SYSTEM ImportExportTestSystem (* System with a device and resource *)
  (* Standard: 61499-1; Description: Copyright (c) 2026 Martin Erich Jobst This program and the accompanying materials are made available under the terms of the Eclipse Public License 2.0 which is available at https://www.eclipse.org/legal/epl-2.0/ SPDX-License-Identifier: EPL-2.0 *)
  (* Version 1.0, 2026-10-23, Martin Jobst *)
  {SET_ATTRIBUTE(IntegerAttribute, 18)}
  APPLICATION TestApplication (* Application using the basic FB *)
    {SET_ATTRIBUTE(IntegerAttribute, 19)}
    (* Application network comment *)
    FBS
      Basic : fixture::basic::BasicTest;
      Composite : CompositeTest;
      Mapped : fixture::basic::BasicTest;
      Mapped2 : fixture::basic::BasicTest;
    END_FBS
    EVENT_CONNECTIONS
      Basic.CNF TO Composite.REQ; (* Application event connection *)
      Mapped.CNF TO Mapped2.REQ; (* Mapped event connection *)
    END_CONNECTIONS
    DATA_CONNECTIONS
      Basic.DO1 TO Composite.DI1; {SET_ATTRIBUTE(Negated, TRUE)}
    END_CONNECTIONS
    ADAPTER_CONNECTIONS
      Basic.EVENT TO Composite.EVENT;
    END_CONNECTIONS
  END_APPLICATION
  DEVICE TestDeviceInstance : TestDevice(DEVICE_ID := DINT#17 {SET_ATTRIBUTE(IntegerAttribute, 21)}) (* Fixture device *)
    {SET_ATTRIBUTE(Profile, FixtureProfile)}
    {SET_ATTRIBUTE(IntegerAttribute, 22)}
    RESOURCE TestResourceInstance : TestResource(RESOURCE_ID := DINT#23) (* Fixture resource *)
      {SET_ATTRIBUTE(IntegerAttribute, 23)}
      FBS
        Processor : fixture::basic::BasicTest;
        Controller : CompositeTest;
      END_FBS
      EVENT_CONNECTIONS
        Processor.CNF TO Controller.REQ; (* Resource event connection *)
      END_CONNECTIONS
      DATA_CONNECTIONS
        Processor.DO1 TO Controller.DI1;
      END_CONNECTIONS
      ADAPTER_CONNECTIONS
        Processor.EVENT TO Controller.EVENT;
      END_CONNECTIONS
    END_RESOURCE
  END_DEVICE
  MAPPINGS
    TestApplication.Mapped ON TestDeviceInstance.TestResourceInstance;
    TestApplication.Mapped2 ON TestDeviceInstance.TestResourceInstance;
  END_MAPPINGS
  SEGMENTS
    TestSegmentInstance : TestSegment; (* Fixture segment *) {SET_ATTRIBUTE(IntegerAttribute, 24)}
  END_SEGMENTS
  LINKS
    TestDeviceInstance => TestSegmentInstance; (* Fixture link *)
  END_LINKS
END_SYSTEM
(* other elements stored in the file *)
(* Attribute Name=IntegerAttribute Value=25 *)
